(* IEC 61131-3 sources: plcassist-cli/packages/volt-lsp-iec/test-corpus/bakon-nano/Device/Plc Logic/Application/Library Manager/CAA Storage, 58 files *)

(* ---- CAASTORAGEVERSIONCONSTANTS.gvl ---- *)
VAR_GLOBAL
	_CAASTORAGE_VERSION_LARGEROREQUAL_3_5_5_0_ : INT := 0;
	_CAASTORAGE_VERSION_LARGEROREQUAL_3_5_8_0_ : INT := 0;
	_CAASTORAGE_VERSION_LARGEROREQUAL_3_5_9_0_ : INT := 0;
	_CAASTORAGE_VERSION_LARGEROREQUAL_3_5_11_10_ : INT := 0;
END_VAR

(* ---- VERSIONCONSTANTS.gvl ---- *)
VAR_GLOBAL
	GC_BYVERSION : BYTE := 1;
	GC_BYVERSION_1 : BYTE := 0;
END_VAR

(* ---- ICURSOR.itf ---- *)
INTERFACE ICURSOR
END_INTERFACE

METHOD CURSORCLOSE : ERROR
END_METHOD

METHOD CURSORMOVE : ERROR
VAR_INPUT
	EDIRECTION : DIRECTION;
END_VAR
END_METHOD

METHOD CURSORSEARCHROWID : ERROR
VAR_INPUT
	IDROW : CAA.IDENT;
END_VAR
END_METHOD

METHOD CURSORSEARCH_DINT : ERROR
VAR_INPUT
	DIVALUE : DINT;
END_VAR
END_METHOD

METHOD CURSORSEARCH_INT : ERROR
VAR_INPUT
	IVALUE : INT;
END_VAR
END_METHOD

METHOD CURSORSEARCH_LINT : ERROR
VAR_INPUT
	LIVALUE : LINT;
END_VAR
END_METHOD

METHOD CURSORSEARCH_LREAL : ERROR
VAR_INPUT
	LRVALUE : LREAL;
END_VAR
END_METHOD

METHOD CURSORSEARCH_NULL : ERROR
END_METHOD

METHOD CURSORSEARCH_REAL : ERROR
VAR_INPUT
	RVALUE : REAL;
END_VAR
END_METHOD

METHOD CURSORSEARCH_SINT : ERROR
VAR_INPUT
	SIVALUE : SINT;
END_VAR
END_METHOD

METHOD CURSORSEARCH_TEXT : ERROR
VAR_IN_OUT
	TXTVALUE : TEXT;
END_VAR
END_METHOD

(* ---- ICURSOR2.itf ---- *)
INTERFACE ICURSOR2
END_INTERFACE

METHOD CURSORSEARCHROWID2 : ERROR
VAR_INPUT
	IDROW : LINT;
END_VAR
END_METHOD

(* ---- ICURSOR3.itf ---- *)
INTERFACE ICURSOR3
END_INTERFACE

(* ---- ICURSORASYNC.itf ---- *)
INTERFACE ICURSORASYNC
END_INTERFACE

METHOD CURSORCLOSEASYNC : PROC_STATE
VAR_INPUT
	ECMD : PROC_CMD;
END_VAR
VAR_OUTPUT
	EERROR : ERROR;
END_VAR
END_METHOD

METHOD CURSORMOVEASYNC : PROC_STATE
VAR_INPUT
	ECMD : PROC_CMD;
	EDIRECTION : DIRECTION;
END_VAR
VAR_OUTPUT
	EERROR : ERROR;
END_VAR
END_METHOD

METHOD CURSORSEARCHROWIDASYNC : PROC_STATE
VAR_INPUT
	ECMD : PROC_CMD;
	IDROW : CAA.IDENT;
END_VAR
VAR_OUTPUT
	EERROR : ERROR;
END_VAR
END_METHOD

METHOD CURSORSEARCH_DINTASYNC : PROC_STATE
VAR_INPUT
	ECMD : PROC_CMD;
	DIVALUE : DINT;
END_VAR
VAR_OUTPUT
	EERROR : ERROR;
END_VAR
END_METHOD

METHOD CURSORSEARCH_INTASYNC : PROC_STATE
VAR_INPUT
	ECMD : PROC_CMD;
	IVALUE : INT;
END_VAR
VAR_OUTPUT
	EERROR : ERROR;
END_VAR
END_METHOD

METHOD CURSORSEARCH_LINTASYNC : PROC_STATE
VAR_INPUT
	ECMD : PROC_CMD;
	LIVALUE : LINT;
END_VAR
VAR_OUTPUT
	EERROR : ERROR;
END_VAR
END_METHOD

METHOD CURSORSEARCH_LREALASYNC : PROC_STATE
VAR_INPUT
	ECMD : PROC_CMD;
	LRVALUE : LREAL;
END_VAR
VAR_OUTPUT
	EERROR : ERROR;
END_VAR
END_METHOD

METHOD CURSORSEARCH_NULLASYNC : PROC_STATE
VAR_INPUT
	ECMD : PROC_CMD;
END_VAR
VAR_OUTPUT
	EERROR : ERROR;
END_VAR
END_METHOD

METHOD CURSORSEARCH_REALASYNC : PROC_STATE
VAR_INPUT
	ECMD : PROC_CMD;
	RVALUE : REAL;
END_VAR
VAR_OUTPUT
	EERROR : ERROR;
END_VAR
END_METHOD

METHOD CURSORSEARCH_SINTASYNC : PROC_STATE
VAR_INPUT
	ECMD : PROC_CMD;
	SIVALUE : SINT;
END_VAR
VAR_OUTPUT
	EERROR : ERROR;
END_VAR
END_METHOD

METHOD CURSORSEARCH_TEXTASYNC : PROC_STATE
VAR_INPUT
	ECMD : PROC_CMD;
END_VAR
VAR_OUTPUT
	EERROR : ERROR;
END_VAR
VAR_IN_OUT
	TXTVALUE : TEXT;
END_VAR
END_METHOD

(* ---- IROW.itf ---- *)
INTERFACE IROW
END_INTERFACE

METHOD ROWUPDATE : ERROR
END_METHOD

(* ---- IROW2.itf ---- *)
INTERFACE IROW2
END_INTERFACE

METHOD GETROWID : ERROR
VAR_OUTPUT
	IDROW : LINT;
END_VAR
END_METHOD

(* ---- IROW3.itf ---- *)
INTERFACE IROW3
END_INTERFACE

(* ---- IROWASYNC.itf ---- *)
INTERFACE IROWASYNC
END_INTERFACE

METHOD ROWUPDATEASYNC : PROC_STATE
VAR_INPUT
	ECMD : PROC_CMD;
END_VAR
VAR_OUTPUT
	EERROR : ERROR;
END_VAR
END_METHOD

(* ---- IROWBASE.itf ---- *)
INTERFACE IROWBASE
END_INTERFACE

METHOD COLUMNGETTYPE : COLUMN_TYPE
VAR_INPUT
	IDCOLUMN : CAA.IDENT;
END_VAR
VAR_OUTPUT
	EERROR : ERROR;
END_VAR
END_METHOD

METHOD ROWCLEAR : ERROR
END_METHOD

METHOD ROWRELEASE : ERROR
END_METHOD

METHOD COLUMNGET_BLOB : ERROR
VAR_INPUT
	IDCOLUMN : CAA.IDENT;
END_VAR
VAR_OUTPUT
	XNULL : BOOL;
END_VAR
VAR_IN_OUT
	BLOBVALUE : BLOB;
END_VAR
END_METHOD

METHOD COLUMNGET_DINT : ERROR
VAR_INPUT
	IDCOLUMN : CAA.IDENT;
END_VAR
VAR_OUTPUT
	DIVALUE : DINT;
	XNULL : BOOL;
END_VAR
END_METHOD

METHOD COLUMNGET_INT : ERROR
VAR_INPUT
	IDCOLUMN : CAA.IDENT;
END_VAR
VAR_OUTPUT
	IVALUE : INT;
	XNULL : BOOL;
END_VAR
END_METHOD

METHOD COLUMNGET_LINT : ERROR
VAR_INPUT
	IDCOLUMN : CAA.IDENT;
END_VAR
VAR_OUTPUT
	LIVALUE : LINT;
	XNULL : BOOL;
END_VAR
END_METHOD

METHOD COLUMNGET_LREAL : ERROR
VAR_INPUT
	IDCOLUMN : CAA.IDENT;
END_VAR
VAR_OUTPUT
	LRVALUE : LREAL;
	XNULL : BOOL;
END_VAR
END_METHOD

METHOD COLUMNGET_REAL : ERROR
VAR_INPUT
	IDCOLUMN : CAA.IDENT;
END_VAR
VAR_OUTPUT
	RVALUE : REAL;
	XNULL : BOOL;
END_VAR
END_METHOD

METHOD COLUMNGET_SINT : ERROR
VAR_INPUT
	IDCOLUMN : CAA.IDENT;
END_VAR
VAR_OUTPUT
	SIVALUE : SINT;
	XNULL : BOOL;
END_VAR
END_METHOD

METHOD COLUMNGET_TEXT : ERROR
VAR_INPUT
	IDCOLUMN : CAA.IDENT;
END_VAR
VAR_OUTPUT
	XNULL : BOOL;
END_VAR
VAR_IN_OUT
	TXTVALUE : TEXT;
END_VAR
END_METHOD

METHOD COLUMNSET_BLOB : ERROR
VAR_INPUT
	IDCOLUMN : CAA.IDENT;
END_VAR
VAR_IN_OUT
	BLOBVALUE : BLOB;
END_VAR
END_METHOD

METHOD COLUMNSET_DINT : ERROR
VAR_INPUT
	IDCOLUMN : CAA.IDENT;
	DIVALUE : DINT;
END_VAR
END_METHOD

METHOD COLUMNSET_INT : ERROR
VAR_INPUT
	IDCOLUMN : CAA.IDENT;
	IVALUE : INT;
END_VAR
END_METHOD

METHOD COLUMNSET_LINT : ERROR
VAR_INPUT
	IDCOLUMN : CAA.IDENT;
	LIVALUE : LINT;
END_VAR
END_METHOD

METHOD COLUMNSET_LREAL : ERROR
VAR_INPUT
	IDCOLUMN : CAA.IDENT;
	LRVALUE : LREAL;
END_VAR
END_METHOD

METHOD COLUMNSET_NULL : ERROR
VAR_INPUT
	IDCOLUMN : CAA.IDENT;
END_VAR
END_METHOD

METHOD COLUMNSET_REAL : ERROR
VAR_INPUT
	IDCOLUMN : CAA.IDENT;
	RVALUE : REAL;
END_VAR
END_METHOD

METHOD COLUMNSET_SINT : ERROR
VAR_INPUT
	IDCOLUMN : CAA.IDENT;
	SIVALUE : SINT;
END_VAR
END_METHOD

METHOD COLUMNSET_TEXT : ERROR
VAR_INPUT
	IDCOLUMN : CAA.IDENT;
END_VAR
VAR_IN_OUT
	TXTVALUE : TEXT;
END_VAR
END_METHOD

METHOD COLUMNUPDATE_BLOB : ERROR
VAR_INPUT
	IDCOLUMN : CAA.IDENT;
END_VAR
VAR_IN_OUT
	BLOBVALUE : BLOB;
	XNULL : BOOL;
END_VAR
END_METHOD

METHOD COLUMNUPDATE_DINT : ERROR
VAR_INPUT
	IDCOLUMN : CAA.IDENT;
END_VAR
VAR_IN_OUT
	DIVALUE : DINT;
	XNULL : BOOL;
END_VAR
END_METHOD

METHOD COLUMNUPDATE_INT : ERROR
VAR_INPUT
	IDCOLUMN : CAA.IDENT;
END_VAR
VAR_IN_OUT
	IVALUE : INT;
	XNULL : BOOL;
END_VAR
END_METHOD

METHOD COLUMNUPDATE_LINT : ERROR
VAR_INPUT
	IDCOLUMN : CAA.IDENT;
END_VAR
VAR_IN_OUT
	LIVALUE : LINT;
	XNULL : BOOL;
END_VAR
END_METHOD

METHOD COLUMNUPDATE_LREAL : ERROR
VAR_INPUT
	IDCOLUMN : CAA.IDENT;
END_VAR
VAR_IN_OUT
	LRVALUE : LREAL;
	XNULL : BOOL;
END_VAR
END_METHOD

METHOD COLUMNUPDATE_REAL : ERROR
VAR_INPUT
	IDCOLUMN : CAA.IDENT;
END_VAR
VAR_IN_OUT
	RVALUE : REAL;
	XNULL : BOOL;
END_VAR
END_METHOD

METHOD COLUMNUPDATE_SINT : ERROR
VAR_INPUT
	IDCOLUMN : CAA.IDENT;
END_VAR
VAR_IN_OUT
	SIVALUE : SINT;
	XNULL : BOOL;
END_VAR
END_METHOD

METHOD COLUMNUPDATE_TEXT : ERROR
VAR_INPUT
	IDCOLUMN : CAA.IDENT;
END_VAR
VAR_IN_OUT
	TXTVALUE : TEXT;
	XNULL : BOOL;
END_VAR
END_METHOD

(* ---- IROWPLANCHET.itf ---- *)
INTERFACE IROWPLANCHET
END_INTERFACE

METHOD ROWINSERT : CAA.IDENT
VAR_OUTPUT
	EERROR : ERROR;
END_VAR
END_METHOD

(* ---- IROWPLANCHETASYNC.itf ---- *)
INTERFACE IROWPLANCHETASYNC
END_INTERFACE

METHOD ROWINSERTASYNC : PROC_STATE
VAR_INPUT
	ECMD : PROC_CMD;
END_VAR
VAR_OUTPUT
	EERROR : ERROR;
END_VAR
END_METHOD

(* ---- ISAVEPOINT.itf ---- *)
INTERFACE ISAVEPOINT
END_INTERFACE

METHOD SAVEPOINTRELEASE : ERROR
END_METHOD

METHOD SAVEPOINTROLLBACK : ERROR
END_METHOD

(* ---- ISAVEPOINTASYNC.itf ---- *)
INTERFACE ISAVEPOINTASYNC
END_INTERFACE

METHOD SAVEPOINTRELEASEASYNC : PROC_STATE
VAR_INPUT
	ECMD : PROC_CMD;
END_VAR
VAR_OUTPUT
	EERROR : ERROR;
END_VAR
END_METHOD

METHOD SAVEPOINTROLLBACKASYNC : PROC_STATE
VAR_INPUT
	ECMD : PROC_CMD;
END_VAR
VAR_OUTPUT
	EERROR : ERROR;
END_VAR
END_METHOD

(* ---- ISTORAGE.itf ---- *)
INTERFACE ISTORAGE
END_INTERFACE

METHOD STORAGECLEAR : ERROR
END_METHOD

METHOD STORAGECLOSE : ERROR
END_METHOD

METHOD STORAGEGETMETRICS : ERROR
VAR_IN_OUT
	MMETRICS : METRICS;
END_VAR
END_METHOD

METHOD STORAGEGETPATH : ERROR
VAR_IN_OUT
	SPATH : CAA.FILENAME;
END_VAR
END_METHOD

METHOD STORAGEOPENFILE : ERROR
VAR_INPUT
	XREADONLY : BOOL;
END_VAR
VAR_IN_OUT
	SPATH : CAA.FILENAME;
END_VAR
END_METHOD

METHOD STORAGEREORG : ERROR
END_METHOD

METHOD TABLEOPEN : ITable
VAR_INPUT
	IDTABLE : CAA.IDENT;
END_VAR
VAR_OUTPUT
	EERROR : ERROR;
END_VAR
END_METHOD

METHOD TRANSACTIONBEGIN : ITransaction
VAR_INPUT
	EMODE : TRANSACTION_MODE;
END_VAR
VAR_OUTPUT
	EERROR : ERROR;
END_VAR
END_METHOD

METHOD UTILITYGETCURRENTDATEANDTIME : INT64
VAR_OUTPUT
	EERROR : ERROR;
END_VAR
END_METHOD

METHOD UTILITYRANDOMNESS : ERROR
VAR_INPUT
	SZSIZE : CAA.SIZE;
	PDATA : CAA.PVOID;
END_VAR
END_METHOD

(* ---- ISTORAGE2.itf ---- *)
INTERFACE ISTORAGE2
END_INTERFACE

METHOD STORAGEEXECUTESTATEMENT : ERROR
VAR_IN_OUT
	SSTATEMENT : SQLSTATEMENT;
END_VAR
END_METHOD

METHOD STORAGEGETINDEXID : ERROR
VAR_OUTPUT
	IDINDEX : CAA.IDENT;
END_VAR
VAR_IN_OUT
	SINDEX : STRING;
	STABLE : STRING;
END_VAR
END_METHOD

METHOD STORAGEGETTABLEID : ERROR
VAR_OUTPUT
	IDTABLE : CAA.IDENT;
END_VAR
VAR_IN_OUT
	STABLE : STRING;
END_VAR
END_METHOD

(* ---- ISTORAGEASYNC.itf ---- *)
INTERFACE ISTORAGEASYNC
END_INTERFACE

METHOD STORAGECLEARASYNC : PROC_STATE
VAR_INPUT
	ECMD : PROC_CMD;
END_VAR
VAR_OUTPUT
	EERROR : ERROR;
END_VAR
END_METHOD

METHOD STORAGECLOSEASYNC : PROC_STATE
VAR_INPUT
	ECMD : PROC_CMD;
END_VAR
VAR_OUTPUT
	EERROR : ERROR;
END_VAR
END_METHOD

METHOD STORAGEOPENFILEASYNC : PROC_STATE
VAR_INPUT
	ECMD : PROC_CMD;
	XREADONLY : BOOL := FALSE;
END_VAR
VAR_OUTPUT
	EERROR : ERROR;
END_VAR
VAR_IN_OUT
	SPATH : CAA.FILENAME;
	ITFSTORAGE : IStorage;
END_VAR
END_METHOD

METHOD STORAGEREORGASYNC : PROC_STATE
VAR_INPUT
	ECMD : PROC_CMD;
END_VAR
VAR_OUTPUT
	EERROR : ERROR;
END_VAR
END_METHOD

METHOD TABLEOPENASYNC : PROC_STATE
VAR_INPUT
	ECMD : PROC_CMD;
	IDTABLE : CAA.IDENT;
END_VAR
VAR_OUTPUT
	ITFTABLE : ITable;
	EERROR : ERROR;
END_VAR
END_METHOD

METHOD TRANSACTIONBEGINASYNC : PROC_STATE
VAR_INPUT
	ECMD : PROC_CMD;
	EMODE : TRANSACTION_MODE;
END_VAR
VAR_OUTPUT
	ITFTRANSACTION : ITransaction;
	EERROR : ERROR;
END_VAR
END_METHOD

(* ---- ITABLE.itf ---- *)
INTERFACE ITABLE
END_INTERFACE

METHOD CURSOROPEN : ICursor
VAR_INPUT
	IDINDEX : CAA.IDENT;
	XREADONLY : BOOL;
END_VAR
VAR_OUTPUT
	EERROR : ERROR;
END_VAR
END_METHOD

METHOD ROWCREATE : IRowPlanchet
VAR_OUTPUT
	EERROR : ERROR;
END_VAR
END_METHOD

METHOD ROWDELETE : ERROR
VAR_INPUT
	IDROW : CAA.IDENT;
END_VAR
END_METHOD

METHOD ROWDUPLICATE : IRowPlanchet
VAR_INPUT
	IDROW : CAA.IDENT;
END_VAR
VAR_OUTPUT
	EERROR : ERROR;
END_VAR
END_METHOD

METHOD ROWSELECT : IRow
VAR_INPUT
	IDROW : CAA.IDENT;
END_VAR
VAR_OUTPUT
	EERROR : ERROR;
END_VAR
END_METHOD

METHOD TABLECLEAR : ERROR
END_METHOD

METHOD TABLECLOSE : ERROR
END_METHOD

(* ---- ITABLE2.itf ---- *)
INTERFACE ITABLE2
END_INTERFACE

METHOD ROWDELETE2 : ERROR
VAR_INPUT
	IDROW : LINT;
END_VAR
END_METHOD

(* ---- ITABLE3.itf ---- *)
INTERFACE ITABLE3
END_INTERFACE

(* ---- ITABLE4.itf ---- *)
INTERFACE ITABLE4
END_INTERFACE

METHOD GETMINMAXROWIDS : ERROR
VAR_OUTPUT
	IDROWMIN : LINT;
	IDROWMAX : LINT;
END_VAR
END_METHOD

(* ---- ITABLEASYNC.itf ---- *)
INTERFACE ITABLEASYNC
END_INTERFACE

METHOD CURSOROPENASYNC : PROC_STATE
VAR_INPUT
	ECMD : PROC_CMD;
	IDCURSOR : CAA.IDENT;
	XREADONLY : BOOL;
END_VAR
VAR_OUTPUT
	ITFCURSOR : ICursor;
	EERROR : ERROR;
END_VAR
END_METHOD

METHOD ROWDELETEASYNC : PROC_STATE
VAR_INPUT
	ECMD : PROC_CMD;
	IDROW : CAA.IDENT;
END_VAR
VAR_OUTPUT
	EERROR : ERROR;
END_VAR
END_METHOD

METHOD ROWSELECTASYNC : PROC_STATE
VAR_INPUT
	ECMD : PROC_CMD;
	IDROW : CAA.IDENT;
END_VAR
VAR_OUTPUT
	ITFROW : IRow;
	EERROR : ERROR;
END_VAR
END_METHOD

METHOD TABLECLEARASYNC : PROC_STATE
VAR_INPUT
	ECMD : PROC_CMD;
END_VAR
VAR_OUTPUT
	EERROR : ERROR;
END_VAR
END_METHOD

METHOD TABLECLOSEASYNC : PROC_STATE
VAR_INPUT
	ECMD : PROC_CMD;
END_VAR
VAR_OUTPUT
	EERROR : ERROR;
END_VAR
END_METHOD

(* ---- ITRANSACTION.itf ---- *)
INTERFACE ITRANSACTION
END_INTERFACE

METHOD TRANSACTIONSETSAVEPOINT : ISavepoint
VAR_OUTPUT
	EERROR : ERROR;
END_VAR
END_METHOD

METHOD TRANSACTIONCOMMIT : ERROR
END_METHOD

METHOD TRANSACTIONROLLBACK : ERROR
END_METHOD

(* ---- ITRANSACTIONASYNC.itf ---- *)
INTERFACE ITRANSACTIONASYNC
END_INTERFACE

METHOD TRANSACTIONSETSAVEPOINTASYNC : PROC_STATE
VAR_INPUT
	ECMD : PROC_CMD;
END_VAR
VAR_OUTPUT
	ITFSAVEPOINT : ISavepoint;
	EERROR : ERROR;
END_VAR
END_METHOD

METHOD TRANSACTIONCOMMITASYNC : PROC_STATE
VAR_INPUT
	ECMD : PROC_CMD;
END_VAR
VAR_OUTPUT
	EERROR : ERROR;
END_VAR
END_METHOD

METHOD TRANSACTIONROLLBACKASYNC : PROC_STATE
VAR_INPUT
	ECMD : PROC_CMD;
END_VAR
VAR_OUTPUT
	EERROR : ERROR;
END_VAR
END_METHOD

(* ---- BLOBALLOC.fun ---- *)
FUNCTION BLOBALLOC : POINTER TO STO_BLOB
VAR_INPUT
	SZDATA : CAA.SIZE;
END_VAR
VAR_OUTPUT
	EERROR : ERROR;
END_VAR
END_FUNCTION

(* ---- BLOBCOPYTODATA.fun ---- *)
FUNCTION BLOBCOPYTODATA : ERROR
VAR_INPUT
	PBLOB : POINTER TO STO_BLOB;
	PDATA : POINTER TO BYTE;
	SZDATA : CAA.SIZE;
END_VAR
END_FUNCTION

(* ---- BLOBFREE.fun ---- *)
FUNCTION BLOBFREE : ERROR
VAR_INPUT
	PBLOB : POINTER TO STO_BLOB;
END_VAR
END_FUNCTION

(* ---- CREATETEXTFROMSTRING.fun ---- *)
FUNCTION CREATETEXTFROMSTRING : ERROR
VAR_IN_OUT
	SVALUE : STRING(1);
	TXTVALUE : STO_TEXT;
END_VAR
END_FUNCTION

(* ---- CREATETEXTFROMWSTRING.fun ---- *)
FUNCTION CREATETEXTFROMWSTRING : ERROR
VAR_IN_OUT
	WSVALUE : WSTRING(1);
	TXTVALUE : STO_TEXT;
END_VAR
END_FUNCTION

(* ---- DATACOPYTOBLOB.fun ---- *)
FUNCTION DATACOPYTOBLOB : ERROR
VAR_INPUT
	PDATA : POINTER TO BYTE;
	SZDATA : CAA.SIZE;
	PBLOB : POINTER TO STO_BLOB;
END_VAR
END_FUNCTION

(* ---- DT_TO_INT64.fun ---- *)
FUNCTION DT_TO_INT64 : ERROR
VAR_INPUT
	DTVALUE : DATE_AND_TIME;
END_VAR
VAR_OUTPUT
	I64VALUE : INT64;
END_VAR
END_FUNCTION

(* ---- DT_TO_ISO8601.fun ---- *)
FUNCTION DT_TO_ISO8601 : ERROR
VAR_INPUT
	DTVALUE : DATE_AND_TIME;
END_VAR
VAR_IN_OUT
	SVALUE : ISO8601;
END_VAR
END_FUNCTION

(* ---- DT_TO_REAL8.fun ---- *)
FUNCTION DT_TO_REAL8 : ERROR
VAR_INPUT
	DTVALUE : DATE_AND_TIME;
END_VAR
VAR_OUTPUT
	R8VALUE : REAL8;
END_VAR
END_FUNCTION

(* ---- GETSUPPLIERVERSION.fun ---- *)
FUNCTION GETSUPPLIERVERSION : WORD
VAR_INPUT
	XDUMMY : BOOL;
END_VAR
END_FUNCTION

(* ---- INT64_TO_DT.fun ---- *)
FUNCTION INT64_TO_DT : ERROR
VAR_INPUT
	I64VALUE : INT64;
END_VAR
VAR_OUTPUT
	DTVALUE : DATE_AND_TIME;
END_VAR
END_FUNCTION

(* ---- INT64_TO_ISO8601.fun ---- *)
FUNCTION INT64_TO_ISO8601 : ERROR
VAR_INPUT
	I64VALUE : INT64;
END_VAR
VAR_IN_OUT
	SVALUE : ISO8601;
END_VAR
END_FUNCTION

(* ---- INT64_TO_LOCALTIME.fun ---- *)
FUNCTION INT64_TO_LOCALTIME : ERROR
VAR_INPUT
	I64UTC : INT64;
END_VAR
VAR_OUTPUT
	I64LOCAL : INT64;
END_VAR
END_FUNCTION

(* ---- INT64_TO_LTIME.fun ---- *)
FUNCTION INT64_TO_LTIME : ERROR
VAR_INPUT
	I64VALUE : INT64;
END_VAR
VAR_OUTPUT
	LTVALUE : LTIME;
END_VAR
END_FUNCTION

(* ---- INT64_TO_REAL8.fun ---- *)
FUNCTION INT64_TO_REAL8 : ERROR
VAR_INPUT
	I64VALUE : INT64;
END_VAR
VAR_OUTPUT
	R8VALUE : REAL8;
END_VAR
END_FUNCTION

(* ---- INT64_TO_TIME.fun ---- *)
FUNCTION INT64_TO_TIME : ERROR
VAR_INPUT
	I64VALUE : INT64;
END_VAR
VAR_OUTPUT
	TVALUE : TIME;
END_VAR
END_FUNCTION

(* ---- INT64_TO_UTC.fun ---- *)
FUNCTION INT64_TO_UTC : ERROR
VAR_INPUT
	I64LOCAL : INT64;
END_VAR
VAR_OUTPUT
	I64UTC : INT64;
END_VAR
END_FUNCTION

(* ---- ISO8601_TO_DT.fun ---- *)
FUNCTION ISO8601_TO_DT : ERROR
VAR_OUTPUT
	DTVALUE : DATE_AND_TIME;
END_VAR
VAR_IN_OUT
	SVALUE : ISO8601;
END_VAR
END_FUNCTION

(* ---- ISO8601_TO_LTIME.fun ---- *)
FUNCTION ISO8601_TO_LTIME : ERROR
VAR_OUTPUT
	LTVALUE : LTIME;
END_VAR
VAR_IN_OUT
	SVALUE : ISO8601;
END_VAR
END_FUNCTION

(* ---- ISO8601_TO_TIME.fun ---- *)
FUNCTION ISO8601_TO_TIME : ERROR
VAR_OUTPUT
	TVALUE : TIME;
END_VAR
VAR_IN_OUT
	SVALUE : ISO8601;
END_VAR
END_FUNCTION

(* ---- LTIME_TO_INT64.fun ---- *)
FUNCTION LTIME_TO_INT64 : ERROR
VAR_INPUT
	LTVALUE : LTIME;
END_VAR
VAR_OUTPUT
	I64VALUE : INT64;
END_VAR
END_FUNCTION

(* ---- LTIME_TO_ISO8601.fun ---- *)
FUNCTION LTIME_TO_ISO8601 : ERROR
VAR_INPUT
	LTVALUE : LTIME;
END_VAR
VAR_IN_OUT
	SVALUE : ISO8601;
END_VAR
END_FUNCTION

(* ---- LTIME_TO_REAL8.fun ---- *)
FUNCTION LTIME_TO_REAL8 : ERROR
VAR_INPUT
	LTVALUE : LTIME;
END_VAR
VAR_OUTPUT
	LRVALUE : LREAL;
END_VAR
END_FUNCTION

(* ---- REAL8_TO_DT.fun ---- *)
FUNCTION REAL8_TO_DT : ERROR
VAR_INPUT
	R8VALUE : REAL8;
END_VAR
VAR_OUTPUT
	DTVALUE : DATE_AND_TIME;
END_VAR
END_FUNCTION

(* ---- REAL8_TO_LTIME.fun ---- *)
FUNCTION REAL8_TO_LTIME : ERROR
VAR_INPUT
	R8VALUE : REAL8;
END_VAR
VAR_OUTPUT
	LTVALUE : LTIME;
END_VAR
END_FUNCTION

(* ---- REAL8_TO_TIME.fun ---- *)
FUNCTION REAL8_TO_TIME : ERROR
VAR_INPUT
	R8VALUE : REAL8;
END_VAR
VAR_OUTPUT
	TVALUE : TIME;
END_VAR
END_FUNCTION

(* ---- STORAGEDELETEFILE.fun ---- *)
FUNCTION STORAGEDELETEFILE : ERROR
VAR_IN_OUT
	SPATH : CAA.FILENAME;
END_VAR
END_FUNCTION

(* ---- TEXTCOPYTOSTRING.fun ---- *)
FUNCTION TEXTCOPYTOSTRING : ERROR
VAR_INPUT
	XFREE : BOOL;
END_VAR
VAR_IN_OUT
	TXTVALUE : STO_TEXT;
	SVALUE : STRING(1);
	SZVALUE : CAA.SIZE;
END_VAR
END_FUNCTION

(* ---- TEXTCOPYTOWSTRING.fun ---- *)
FUNCTION TEXTCOPYTOWSTRING : ERROR
VAR_INPUT
	XFREE : BOOL;
END_VAR
VAR_IN_OUT
	TXTVALUE : STO_TEXT;
	WSVALUE : WSTRING(1);
	SZVALUE : CAA.SIZE;
END_VAR
END_FUNCTION

(* ---- TEXTFREE.fun ---- *)
FUNCTION TEXTFREE : ERROR
VAR_IN_OUT
	TXTVALUE : STO_TEXT;
END_VAR
END_FUNCTION

(* ---- TIME_TO_INT64.fun ---- *)
FUNCTION TIME_TO_INT64 : ERROR
VAR_INPUT
	TVALUE : TIME;
END_VAR
VAR_OUTPUT
	I64VALUE : INT64;
END_VAR
END_FUNCTION

(* ---- TIME_TO_ISO8601.fun ---- *)
FUNCTION TIME_TO_ISO8601 : ERROR
VAR_INPUT
	TVALUE : TIME;
END_VAR
VAR_IN_OUT
	SVALUE : ISO8601;
END_VAR
END_FUNCTION

(* ---- TIME_TO_REAL8.fun ---- *)
FUNCTION TIME_TO_REAL8 : ERROR
VAR_INPUT
	TVALUE : TIME;
END_VAR
VAR_OUTPUT
	R8VALUE : REAL8;
END_VAR
END_FUNCTION
